// TIA Portal V21 export
// export: Created 2026-11-22T00:27:54.9526895Z, ExportSetting WithDefaults, DisplayName Totally Integrated Automation Portal, DisplayVersion V21 Update 3, DisplayName STEP 7 Professional, DisplayVersion V21 Update 3, DisplayName STEP 7 Safety, DisplayVersion V21, DisplayName Tech WebApplication, DisplayVersion V21, DisplayName WinCC Basic/Comfort/Advanced, DisplayVersion V21 Update 3, DisplayName WinCC Unified, DisplayVersion V21 Update 3
Screen "P_Gauge_3"  1024x768, Number=120
  ScreenLayer "Layer_0"
    Gauge "ShowLimitRanges" at 10,10 size 150x150  CenterSize=0.08, DialSize=0.87, Gradation=10, InnerDialInnerDistance=0.08, InnerDialOuterDistance=0.9, MaximumValue=100, RangeUpper1Start=3.5, RangeUpper2Start=70, StyleItem=Gauge, CaptionText="SIMATIC"
    TextField "Label_ShowLimitRanges" at 10,162 size 158x16  StyleItem=Text field, Text="ShowLimitRanges"
    Gauge "ShowPeakValuePointer" at 170,10 size 150x150  CenterSize=0.08, DialSize=0.87, Gradation=10, InnerDialInnerDistance=0.08, InnerDialOuterDistance=0.9, MaximumValue=100, RangeUpper1Start=3.5, RangeUpper2Start=70, StyleItem=Gauge, CaptionText="SIMATIC"
    TextField "Label_ShowPeakValuePointer" at 170,162 size 158x16  StyleItem=Text field, Text="ShowPeakValuePointer"
    Gauge "UnitColor" at 330,10 size 150x150  CenterSize=0.08, DialSize=0.87, Gradation=10, InnerDialInnerDistance=0.08, InnerDialOuterDistance=0.9, MaximumValue=100, RangeUpper1Start=3.5, RangeUpper2Start=70, StyleItem=Gauge, CaptionText="SIMATIC"
    TextField "Label_UnitColor" at 330,162 size 158x16  StyleItem=Text field, Text="UnitColor"
    Gauge "UnitTop" at 490,10 size 150x150  CenterSize=0.08, DialSize=0.87, Gradation=10, InnerDialInnerDistance=0.08, InnerDialOuterDistance=0.9, MaximumValue=100, RangeUpper1Start=3.5, RangeUpper2Start=70, StyleItem=Gauge, CaptionText="SIMATIC"
    TextField "Label_UnitTop" at 490,162 size 158x16  StyleItem=Text field, Text="UnitTop"
    Gauge "UseDesignColorSchema" at 650,10 size 150x150  CenterSize=0.08, DialSize=0.87, Gradation=10, InnerDialInnerDistance=0.08, InnerDialOuterDistance=0.9, MaximumValue=100, RangeUpper1Start=3.5, RangeUpper2Start=70, CaptionText="SIMATIC"
    TextField "Label_UseDesignColorSchema" at 650,162 size 158x16  StyleItem=Text field, Text="UseDesignColorSchema"
    Button "Next" at 982,744 size 40x22  Mode=Text, StyleItem=Button, TextOff="Text", TextOn="Text"
      on Click: ActivateScreen(Screen name := P_Clock_1, Object number := 0)
